(* IEC 61131-3 sources: verifaps-lib/util/src/testFixtures/resources/edu/kit/iti/formal/automation/st/types, 10 files *)

(* ---- array1.st ---- *)
TYPE
    ary : ARRAY[1..10] OF SINT;
    ary : ARRAY[1..10,100..10] OF SINT;
    ary : ARRAY[1..10,-12..12] OF SINT;
//error    ary : ARRAY[1..2] OF ARRAY[1..2];
    ary : ARRAY[1..10,1..1,1..1,1..1,1..1,1..1,1..1,1..1,1..1,1..1,
    1..1,1..1,1..1,1..1,1..1,1..1,1..1,1..1,1..1] OF Blub;
END_TYPE

(* ---- enum_1.st ---- *)
TYPE  MY_ENUM : (one, two, three);
                   END_TYPE

(* ---- struct1.st ---- *)
TYPE
S : STRUCT
    A: INT;
    B: INT:= 3;
    C: BOOL;
END_STRUCT;
END_TYPE

(* ---- types1.st ---- *)
TYPE
    A : INT;
    B : INT := 2;
    C : BOOL;
    D : A;
END_TYPE

(* ---- types_1.st ---- *)
TYPE wochtentag_type : (mon, die, mit , don, fre,sam, son); END_TYPE

(* ---- types_2.st ---- *)
TYPE
        temperatur : INT (-40..70);
        monatstage : INT(1..31);
END_TYPE

(* ---- types_3.st ---- *)
    TYPE feld: ARRAY[1..16] of INT;
END_TYPE

(* ---- types_4.st ---- *)
TYPE
    waehrungs_typ : (Euro,Dollar,Yen,Pfund,Default) := Default;
    //subrange fertigungstage: wochentag_typ (mon..fre);
END_TYPE

(* ---- types_5.st ---- *)
TYPE f: feld;
     i: INTEGER;
END_TYPE

(* ---- types_6.st ---- *)
TYPE temp_sig :
        STRUCT
            temp:temperatur;
            filter_param: SINT (0..99);
        END_STRUCT;
END_TYPE
